{attribute 'qualified_only'}
{attribute 'strict'}
{attribute 'to_string'}
TYPE E_IdGenFailureReason :
(
	NA := 0,  // No failure occurred.
	NO_IDENTIFIERS_AVAILABLE,  // The ring held too few bytes; the caller must retry on a later cycle.
	GUID_SERVICE_FAILED,  // The TwinCAT GUID service reported an error while the ring was being refilled.
	MEMORY_ALLOCATION_FAILURE,  // The ring could not be allocated.
	INVALID_CONFIGUATION  // parameters used to configure the generator were not valid
) UDINT;
END_TYPE

(* stored: Version 1.1.0.1
   EnumerationTextList E_IdGenFailureReason: Id {9278004f-779f-4ad2-a921-a0e4dfcd69b1} *)
